ABB RAPID module: ConfProg.mod

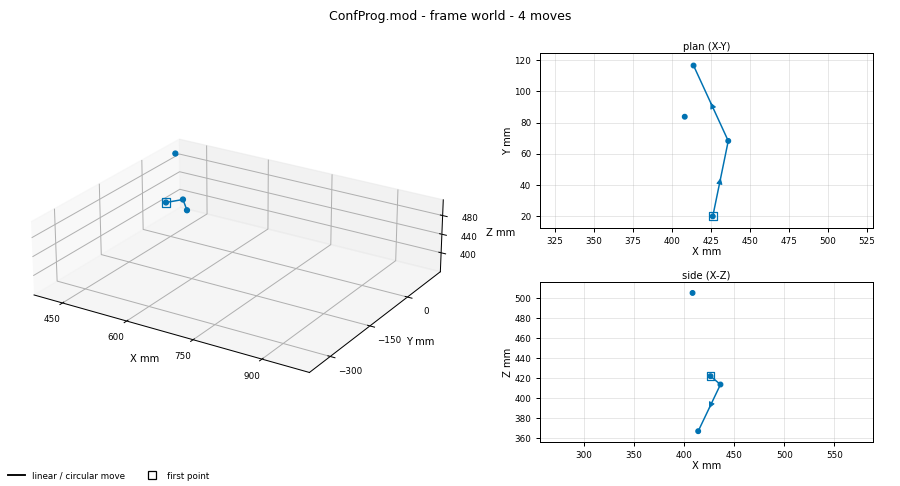
[picture p0: tool path of ConfProg.mod in frame world, 4 of 6 moves have a stored position in this frame; points joined in program order, loops and branches not executed]
%%%
  VERSION:1
  LANGUAGE:ENGLISH
%%%
MODULE MOD_ConfProg

    ! -------------------------------
    ! Define customized variables here
    ! ...

	! Tool variables:
	PERS tooldata ToolS := [TRUE,[[10.000,20.000,150.000],[1.00000000,0.00000000,0.00000000,0.00000000]],[1,[0,0,20],[1,0,0,0],0,0,0.005]];

	! Reference variables:
	PERS wobjdata FrameS := [FALSE, TRUE, "", [[0,0,0],[1,0,0,0]],[[1234.570,-98.765,50.500],[0.96592583,0.00000000,0.00000000,0.25881905]]];

	PROC Main()
		ConfJ \On;
		ConfL \Off;
		! Program generated by RoboDK v6.0.7 for ABB IRB 260 on XX/XX/XXXX 18:00:00
		! Using nominal kinematics.
		MoveL [[-640.584,506.980,371.534],[0.37410804,0.28584607,0.85365954,-0.22271191],[0,0,0,0],[9E+09,9E+09,9E+09,9E+09,9E+09,9E+09]],v500,z1,ToolS \WObj:=FrameS;
		MoveL [[-607.850,543.849,363.215],[0.37410804,0.28584607,0.85365954,-0.22271191],[0,0,0,4],[9E+09,9E+09,9E+09,9E+09,9E+09,9E+09]],v500,z1,ToolS \WObj:=FrameS;
		MoveL [[-602.951,596.788,316.595],[0.37410804,0.28584607,0.85365954,-0.22271191],[0,0,0,3],[9E+09,9E+09,9E+09,9E+09,9E+09,9E+09]],v500,z1,ToolS \WObj:=FrameS;
		MoveAbsJ [[10.000000,20.000000,-30.000000,40.000000,0.000000,0.000000],[9E+09,9E+09,9E+09,9E+09,9E+09,9E+09]],v500,z1,ToolS \WObj:=FrameS;
		MoveAbsJ [[-170.000000,45.000000,-45.000000,-170.000000,0.000000,0.000000],[9E+09,9E+09,9E+09,9E+09,9E+09,9E+09]],v500,z1,ToolS \WObj:=FrameS;
		MoveC [[-353.026,-90.135,331.702],[0.34432926,0.04805561,0.93307257,-0.09221494],[0,0,0,1],[9E+09,9E+09,9E+09,9E+09,9E+09,9E+09]],[[-624.230,571.208,454.620],[0.55239178,-0.04267608,0.67304167,-0.48995609],[0,0,0,4],[9E+09,9E+09,9E+09,9E+09,9E+09,9E+09]],v500,z1,ToolS \WObj:=FrameS;
	ENDPROC

ENDMODULE
